(* IEC 61131-3 sources: codesys-to-s7/tests/corpus/C2S7-TYPE-ALIAS/neg, 1 file *)

(* ---- input.st ---- *)
TYPE ST_Pct : STRUCT v : INT; END_STRUCT END_TYPE
FUNCTION_BLOCK FB_Case
VAR
    p : ST_Pct;
END_VAR
p.v := 5;
END_FUNCTION_BLOCK
